(*~
	<docu>
		<summary>
			Test type parameter value (code x1000) to test type.
		</summary>
	</docu>
~*)
FUNCTION TcoAteqG6_ToTestType_v_3_5_x : eTcoAteqG6_TestType_v_3_5_x
VAR_INPUT
	inRaw : DINT;
END_VAR

CASE inRaw OF
	0: TcoAteqG6_ToTestType_v_3_5_x := eTcoAteqG6_TestType_v_3_5_x.Invalid;
	1000: TcoAteqG6_ToTestType_v_3_5_x := eTcoAteqG6_TestType_v_3_5_x.Direct;
	2000: TcoAteqG6_ToTestType_v_3_5_x := eTcoAteqG6_TestType_v_3_5_x.Operator;
ELSE
	TcoAteqG6_ToTestType_v_3_5_x := eTcoAteqG6_TestType_v_3_5_x.Unknown;
END_CASE

END_FUNCTION

(* stored: Version 1.1.0.1, ProductVersion 3.1.4024.12
   POU TcoAteqG6_ToTestType_v_3_5_x: Id {8c99c010-77c1-4953-b11c-16d230775a77}, SpecialFunc None *)
